Fanuc KAREL source: KO00044.KL

PROGRAM KO00044
%NOLOCKGROUP
%ENVIRONMENT MIR
VAR
  P1: POSITION
  P2: XYZWPREXT
  F: BOOLEAN
  OUT: JOINTPOS
BEGIN
  F = TRUE
  OUT = MIRROR(P1, P2, F)
END KO00044
